Staubli VAL3: bind.pgx

program bind()
begin
  userPageBindClick("message","btnback",bBack,true)
  userPageBind("message","lst1","options",sRobotMsg,size(sRobotMsg),"r")
end
